// TIA Portal V20 export
// export: Created 2026-10-12T16:46:22.8333962Z, ExportSetting WithDefaults, DisplayName Totally Integrated Automation Portal, DisplayVersion V20 Update 6, DisplayName TIA Portal Openness, DisplayVersion V20 Update 6, DisplayName TIA Portal Version Control Interface, DisplayVersion V20 Update 6, DisplayName SINAMICS Startdrive Advanced, DisplayVersion V20 SP1 Update 2, DisplayName SINAMICS Startdrive G110M, G120, G120C, G120D, G120P, G115D, DisplayVersion V20 SP1 Update 2, DisplayName SINAMICS Startdrive G130, G150, S120, S150, SINAMICS MV, G220, S200, S210, DisplayVersion V20 SP1 Update 2, DisplayName STEP 7 Professional, DisplayVersion V20 Update 6, DisplayName STEP 7 Safety, DisplayVersion V20 Update 2, DisplayName WinCC Basic/Comfort/Advanced, DisplayVersion V20 Update 6, DisplayName WinCC Professional, DisplayVersion V20 Update 6, DisplayName WinCC Unified, DisplayVersion V20 Update 6
TYPE "UDT_WT_Rueckmeldung"
// stored: IsFailsafeCompliant false
   STRUCT
      Belegt : Bool;
      Auftragsindex : Int;
      SchrittIndex : Int;
      Artikel_ID : Int;
      BadNr : Int;
      Personal_ID : Int;
      WT_Eingesetzt : Bool;
      Istzeit : Time;
      Restzeit : Time;
      Verweilzeit_Soll : Time;
      Vorwarn_Erreicht : Bool;
      Zeit_Abgelaufen : Bool;
      Krit_Zeit_Abgelaufen : Bool;
      Stoerung_Aufgetreten : Bool;
      Temp_Abweichung_Max : Real;
      Temp_Toleranz_Eingehalten : Bool;
      Zeitueberschreitung : Time;
      Zeitstempel_Eingesetzt : DTL;
      Zeitstempel_Entnommen : DTL;
      Protokoll_Neu : Bool;
   END_STRUCT;
END_TYPE
